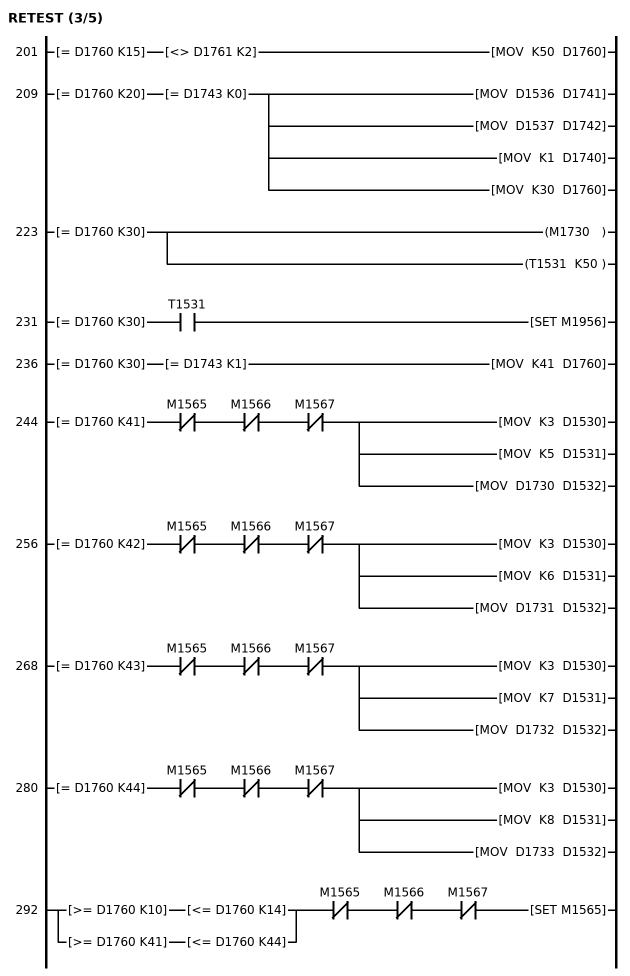
[picture p24: ladder of RETEST, rungs at steps 201 to 292]
201   LD=     D1760 K15
      AND<>   D1761 K2
      MOV     K50 D1760
209   LD=     D1760 K20
      AND=    D1743 K0
      MOV     D1536 D1741
      MOV     D1537 D1742
      MOV     K1 D1740
      MOV     K30 D1760
223   LD=     D1760 K30
      OUT     M1730
      OUT     T1531 K50
231   LD=     D1760 K30
      AND     T1531
      SET     M1956
236   LD=     D1760 K30
      AND=    D1743 K1
      MOV     K41 D1760
244   LD=     D1760 K41
      ANI     M1565
      ANI     M1566
      ANI     M1567
      MOV     K3 D1530
      MOV     K5 D1531
      MOV     D1730 D1532
256   LD=     D1760 K42
      ANI     M1565
      ANI     M1566
      ANI     M1567
      MOV     K3 D1530
      MOV     K6 D1531
      MOV     D1731 D1532
268   LD=     D1760 K43
      ANI     M1565
      ANI     M1566
      ANI     M1567
      MOV     K3 D1530
      MOV     K7 D1531
      MOV     D1732 D1532
280   LD=     D1760 K44
      ANI     M1565
      ANI     M1566
      ANI     M1567
      MOV     K3 D1530
      MOV     K8 D1531
      MOV     D1733 D1532
292   LD>=    D1760 K10
      AND<=   D1760 K14
      LD>=    D1760 K41
      AND<=   D1760 K44
      ORB
      ANI     M1565
      ANI     M1566
      ANI     M1567
      SET     M1565
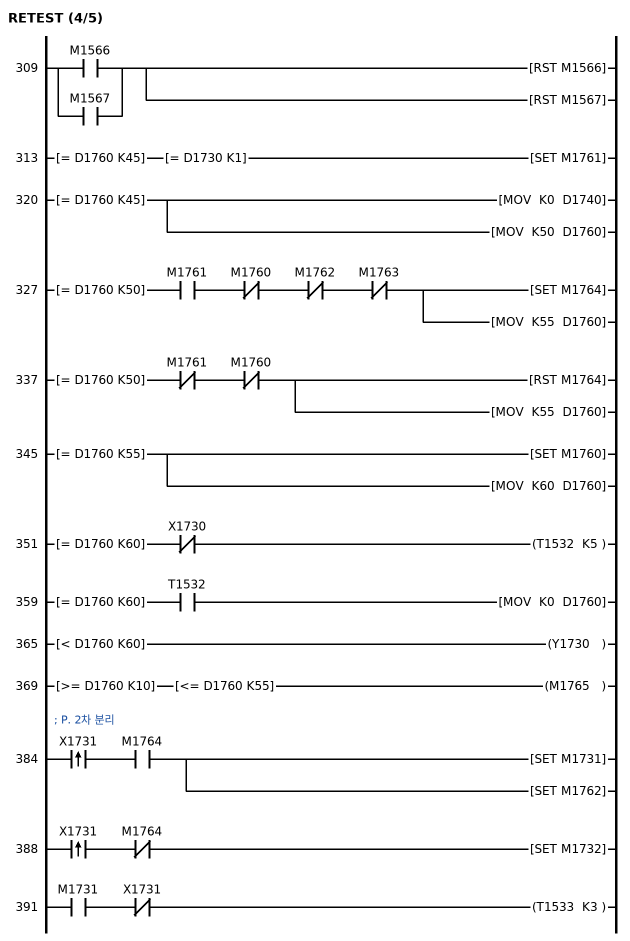
309   LD      M1566
      OR      M1567
      RST     M1566
      RST     M1567
313   LD=     D1760 K45
      AND=    D1730 K1
      SET     M1761
320   LD=     D1760 K45
      MOV     K0 D1740
      MOV     K50 D1760
327   LD=     D1760 K50
      AND     M1761
      ANI     M1760
      ANI     M1762
      ANI     M1763
      SET     M1764
      MOV     K55 D1760
337   LD=     D1760 K50
      ANI     M1761
      ANI     M1760
      RST     M1764
      MOV     K55 D1760
345   LD=     D1760 K55
      SET     M1760
      MOV     K60 D1760
351   LD=     D1760 K60
      ANI     X1730
      OUT     T1532 K5
359   LD=     D1760 K60
      AND     T1532
      MOV     K0 D1760
365   LD<     D1760 K60
      OUT     Y1730
369   LD>=    D1760 K10
      AND<=   D1760 K55
      OUT     M1765
; P. 2차 분리
384   LDP     X1731
      AND     M1764
      SET     M1731
      SET     M1762
388   LDP     X1731
      ANI     M1764
      SET     M1732
391   LD      M1731
      ANI     X1731
      OUT     T1533 K3
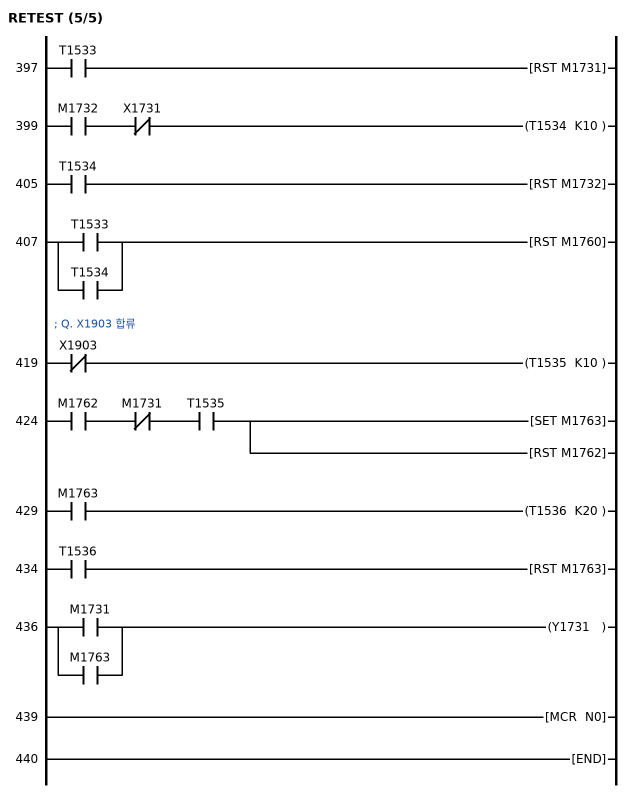
397   LD      T1533
      RST     M1731
399   LD      M1732
      ANI     X1731
      OUT     T1534 K10
405   LD      T1534
      RST     M1732
407   LD      T1533
      OR      T1534
      RST     M1760
; Q. X1903 합류
419   LDI     X1903
      OUT     T1535 K10
424   LD      M1762
      ANI     M1731
      AND     T1535
      SET     M1763
      RST     M1762
429   LD      M1763
      OUT     T1536 K20
434   LD      T1536
      RST     M1763
436   LD      M1731
      OR      M1763
      OUT     Y1731
439   MCR     N0
440   END
END_PROGRAM

PROGRAM DRIVE
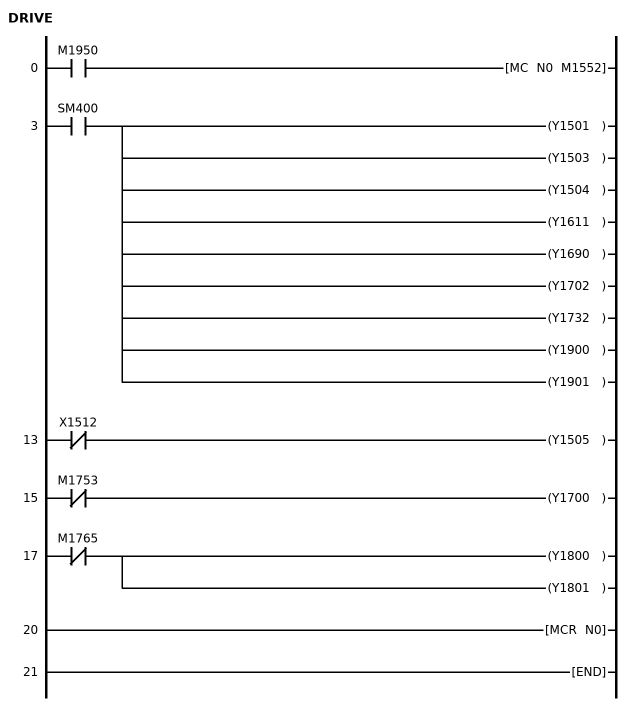
0     LD      M1950
      MC      N0 M1552
3     LD      SM400
      OUT     Y1501
      OUT     Y1503
      OUT     Y1504
      OUT     Y1611
      OUT     Y1690
      OUT     Y1702
      OUT     Y1732
      OUT     Y1900
      OUT     Y1901
13    LDI     X1512
      OUT     Y1505
15    LDI     M1753
      OUT     Y1700
17    LDI     M1765
      OUT     Y1800
      OUT     Y1801
20    MCR     N0
21    END
END_PROGRAM

PROGRAM COUNTER
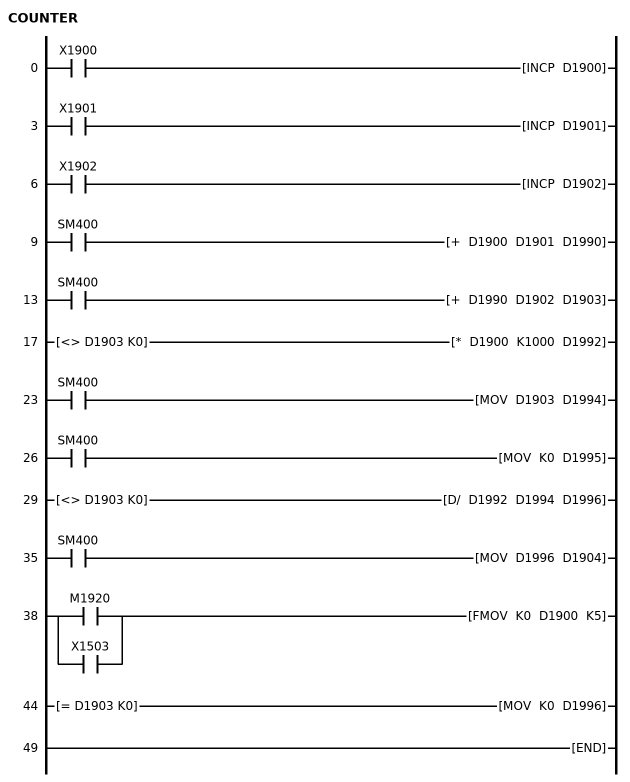
0     LD      X1900
      INCP    D1900
3     LD      X1901
      INCP    D1901
6     LD      X1902
      INCP    D1902
9     LD      SM400
      +       D1900 D1901 D1990
13    LD      SM400
      +       D1990 D1902 D1903
17    LD<>    D1903 K0
      *       D1900 K1000 D1992
23    LD      SM400
      MOV     D1903 D1994
26    LD      SM400
      MOV     K0 D1995
29    LD<>    D1903 K0
      D/      D1992 D1994 D1996
35    LD      SM400
      MOV     D1996 D1904
38    LD      M1920
      OR      X1503
      FMOV    K0 D1900 K5
44    LD=     D1903 K0
      MOV     K0 D1996
49    END
END_PROGRAM

PROGRAM LAMP
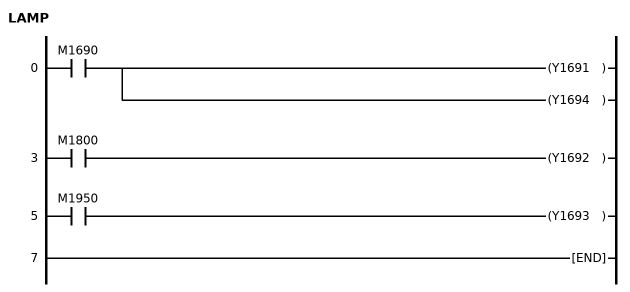
0     LD      M1690
      OUT     Y1691
      OUT     Y1694
3     LD      M1800
      OUT     Y1692
5     LD      M1950
      OUT     Y1693
7     END
END_PROGRAM
